(* IEC 61131-3 sources: Test002/ConveyorBelt/Network, 1 file *)

(* ---- ConfigObjects.st ---- *)
FUNCTION GLOBAL TAB TASK_CONF
_K_TASK, _K_REAL,
_K_END_VAR,

_K_TASK, _K_CYCLIC,
_K_END_VAR,

_K_TASK, _K_BACKGROUND,
_K_END_VAR,

_K_END_CONF
END_FUNCTION

FUNCTION GLOBAL TAB IPR_CONF
_K_IPR
	0$UINT,
_K_END_VAR,
_K_END_CONF
END_FUNCTION

FUNCTION GLOBAL TAB CONFIG_TABLES
00054$UINT,
0$UINT, 0, 4, "_CAN",
0$UINT, 1, 10, "_CANLIB",
0$UINT, 1, 20, "_FILESYS",
0$UINT, 1, 1, "_MULTITASK",
0$UINT, 0, 5, "_OSKERNEL",
0$UINT, 1, 34, "_SERLIB",
0$UINT, 0, 0, "_STDLIB",
0$UINT, 1, 1, "_TASKOBJECTCONTROL",
0$UINT, 1, 18, "AI043",
0$UINT, 1, 20, "ASCII_BIN",
0$UINT, 1, 23, "BUSINTERFACESDIAS",
0$UINT, 2, 0, "BUSINTERFACESDIASINTERNAL",
0$UINT, 1, 0, "CONVEYORBELT",
0$UINT, 1, 1, "CP112_IOS",
0$UINT, 0, 4, "CRITICALSECTION",
0$UINT, 2, 33, "DIASMASTER",
0$UINT, 1, 81, "DIASMASTERC",
0$UINT, 2, 23, "DIASMASTERMAIN",
0$UINT, 1, 0, "DIASMASTERPOSTSCAN",
0$UINT, 1, 13, "DM161",
0$UINT, 1, 11, "EEPROM",
0$UINT, 1, 21, "HUB_BASE",
0$UINT, 2, 11, "HUB_BASE_ROOT",
0$UINT, 2, 35, "HWBASE",
0$UINT, 2, 55, "HWBASECDIAS",
0$UINT, 5, 9, "HWCONTROL",
0$UINT, 1, 10, "HWCONTROLBASE",
0$UINT, 1, 0, "HWRTPOSTSCAN",
0$UINT, 1, 6, "I2CCDIAS",
0$UINT, 1, 22, "MERKEREX",
0$UINT, 1, 9, "RAMFILE",
0$UINT, 1, 20, "SAFETYBASEFSOE",
0$UINT, 3, 16, "SAFETYCDIAS_BASE",
0$UINT, 2, 17, "SAFETYMANAGER",
0$UINT, 1, 3, "SAFETYUDP",
0$UINT, 1, 31, "SCP111",
0$UINT, 1, 59, "SDIASBASE",
0$UINT, 1, 10, "SDIASHUBBASE",
0$UINT, 1, 93, "SDIASMANAGER",
0$UINT, 2, 1, "SDIASPLC",
0$UINT, 1, 9, "SDIASSAFETYBASE",
0$UINT, 1, 23, "SDIASSAFETYMANAGERFSOE",
0$UINT, 1, 10, "SDM081",
0$UINT, 0, 29, "SIGCLIB",
0$UINT, 1, 10, "STRING",
0$UINT, 1, 82, "STRINGINTERNAL",
0$UINT, 1, 21, "SYNCCALL",
0$UINT, 2, 15, "VARAN_BASE",
0$UINT, 3, 2, "VARANMANAGER",
0$UINT, 2, 2, "VARANMANAGER_1",
0$UINT, 1, 24, "VARANMANAGER_BASE",
0$UINT, 1, 3, "VIRTUALBASEINIT",
0$UINT, 2, 11, "WATCHDOGDIAS",
0$UINT, 1, 1, "XXXBASE_IOS",
ONE_CFG$UINT, 0, 0, "ONE_HW_Network",
ONE_CFG$UINT, 0, 0, "ONE_Network0",
TASK_CFG$UINT, 0, 0, "TASK_CONF",
IPR_CFG$UINT, 0, 0, "IPR_CONF",
PRJ_CFG$UINT, 0, 0, "ConveyorBelt",
END_FUNCTION

#ifdef __LSLLDR_IOELEMENTS__
FUNCTION GLOBAL TAB _IO_ELEMENTS_TAB
0001$UINT, 0007$UINT,
"LichtSch01", "DM1611.Input2",
"LichtSch02", "DM1611.Input3",
"Motor01", "DM1611.Output1",
"Motor2", "DM1611.Output3",
"Start01", "DM1611.Input1",
"Zylinder01", "DM1611.Output2",
"Zylinder02", "DM1611.Output4",
0008$UINT,
"LichtSch01", "ConveyorBelt1.Lichtschrank",
"LichtSch01", "ConveyorBelt2.Start",
"LichtSch02", "ConveyorBelt2.Lichtschrank",
"Motor01", "ConveyorBelt1.Motor",
"Motor2", "ConveyorBelt2.Motor",
"Start01", "ConveyorBelt1.Start",
"Zylinder01", "ConveyorBelt1.Cylinder",
"Zylinder02", "ConveyorBelt2.Cylinder",
END_FUNCTION
#endif //__LSLLDR_IOELEMENTS__

FUNCTION GLOBAL TAB CH_REDIRECT_EMB_TAB
0000$UINT,
00014$UINT,
"AI043;SerialNo", "\SerialNoStr.Data",
"BusInterfaceSdias;SerialNo", "\SerialNoStr.Data",
"DM161;SerialNo", "\SerialNoStr.Data",
"HwBaseCDIAS;SerialNo", "\SerialNoStr.Data",
"SCP111;DesignerPrjName", "\SdiasSafetyManagerFSoE1\ProjectNameStr.Data",
"SCP111;DesignerPrjRev", "\SdiasSafetyManagerFSoE1\ProjectRevisionStr.Data",
"SCP111;SerialNo", "\SerialNoStr.Data",
"SDM081;SerialNo", "\SerialNoStr.Data",
"SafetyCDIAS_Base;SerialNo", "\SerialNoStr.Data",
"SdiasBase;SerialNo", "\SerialNoStr.Data",
"SdiasSafetyBase;SerialNo", "\SerialNoStr.Data",
"SdiasSafetyManagerFSoE;DesignerPrjName", "\ProjectNameStr.Data",
"SdiasSafetyManagerFSoE;DesignerPrjRev", "\ProjectRevisionStr.Data",
"Varan_Base;SerialNo", "\SerialNoStr.Data",
END_FUNCTION
